FUNCTION_BLOCK PROCESS_IDENTIFIER (* RLS identification and periodic model-based PID tuning *)
  (* Standard: 61499-2 *)
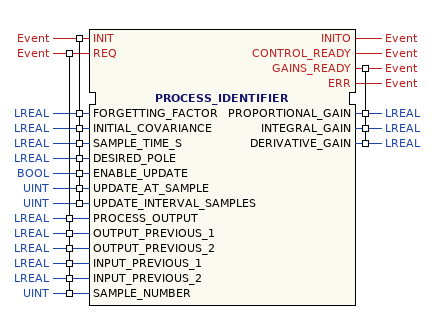
  EVENT_INPUT
    INIT WITH FORGETTING_FACTOR, INITIAL_COVARIANCE, SAMPLE_TIME_S, DESIRED_POLE, ENABLE_UPDATE, UPDATE_AT_SAMPLE, UPDATE_INTERVAL_SAMPLES;
    REQ WITH PROCESS_OUTPUT, OUTPUT_PREVIOUS_1, OUTPUT_PREVIOUS_2, INPUT_PREVIOUS_1, INPUT_PREVIOUS_2, SAMPLE_NUMBER;
  END_EVENT
  EVENT_OUTPUT
    INITO;
    CONTROL_READY;
    GAINS_READY WITH PROPORTIONAL_GAIN, INTEGRAL_GAIN, DERIVATIVE_GAIN;
    ERR;
  END_EVENT
  VAR_INPUT
    FORGETTING_FACTOR : LREAL;
    INITIAL_COVARIANCE : LREAL;
    SAMPLE_TIME_S : LREAL;
    DESIRED_POLE : LREAL;
    ENABLE_UPDATE : BOOL;
    UPDATE_AT_SAMPLE : UINT;
    UPDATE_INTERVAL_SAMPLES : UINT;
    PROCESS_OUTPUT : LREAL;
    OUTPUT_PREVIOUS_1 : LREAL;
    OUTPUT_PREVIOUS_2 : LREAL;
    INPUT_PREVIOUS_1 : LREAL;
    INPUT_PREVIOUS_2 : LREAL;
    SAMPLE_NUMBER : UINT;
  END_VAR
  VAR_OUTPUT
    PROPORTIONAL_GAIN : LREAL;
    INTEGRAL_GAIN : LREAL;
    DERIVATIVE_GAIN : LREAL;
  END_VAR
  FBS
    Estimator : RLS_PARAMETER_ESTIMATOR;
    Trigger : TUNING_TRIGGER;
    Tuner : PID_MODEL_TUNER;
  END_FBS
  EVENT_CONNECTIONS
    INIT TO Estimator.INIT;
    Estimator.INITO TO Trigger.INIT;
    Trigger.INITO TO INITO;
    REQ TO Estimator.REQ;
    Estimator.CNF TO Trigger.REQ;
    Trigger.CONTROL_READY TO CONTROL_READY;
    Trigger.TUNE TO Tuner.REQ;
    Tuner.CNF TO GAINS_READY;
    Estimator.ERR TO ERR;
    Trigger.ERR TO ERR;
    Tuner.ERR TO ERR;
  END_CONNECTIONS
  DATA_CONNECTIONS
    PROCESS_OUTPUT TO Estimator.PROCESS_OUTPUT;
    OUTPUT_PREVIOUS_1 TO Estimator.OUTPUT_PREVIOUS_1;
    OUTPUT_PREVIOUS_2 TO Estimator.OUTPUT_PREVIOUS_2;
    INPUT_PREVIOUS_1 TO Estimator.INPUT_PREVIOUS_1;
    INPUT_PREVIOUS_2 TO Estimator.INPUT_PREVIOUS_2;
    FORGETTING_FACTOR TO Estimator.FORGETTING_FACTOR;
    INITIAL_COVARIANCE TO Estimator.INITIAL_COVARIANCE;
    ENABLE_UPDATE TO Trigger.ENABLE_UPDATE;
    UPDATE_AT_SAMPLE TO Trigger.UPDATE_AT_SAMPLE;
    UPDATE_INTERVAL_SAMPLES TO Trigger.UPDATE_INTERVAL_SAMPLES;
    SAMPLE_NUMBER TO Trigger.SAMPLE_NUMBER;
    SAMPLE_TIME_S TO Tuner.SAMPLE_TIME_S;
    DESIRED_POLE TO Tuner.DESIRED_POLE;
    Estimator.EST_OUTPUT_COEFFICIENT_1 TO Tuner.MODEL_OUTPUT_COEFFICIENT_1;
    Estimator.EST_OUTPUT_COEFFICIENT_2 TO Tuner.MODEL_OUTPUT_COEFFICIENT_2;
    Estimator.EST_INPUT_COEFFICIENT_1 TO Tuner.MODEL_INPUT_COEFFICIENT_1;
    Estimator.EST_INPUT_COEFFICIENT_2 TO Tuner.MODEL_INPUT_COEFFICIENT_2;
    Tuner.TARGET_PROPORTIONAL_GAIN TO PROPORTIONAL_GAIN;
    Tuner.TARGET_INTEGRAL_GAIN TO INTEGRAL_GAIN;
    Tuner.TARGET_DERIVATIVE_GAIN TO DERIVATIVE_GAIN;
  END_CONNECTIONS
END_FUNCTION_BLOCK
